Fanuc KAREL source: KB00181.KL

PROGRAM KB00181
%NOLOCKGROUP
%ENVIRONMENT TIM
VAR
  P1: INTEGER
BEGIN
  P1 = 1
  SET_TIME(P1)
END KB00181
